(*

**Autonumbered labeled footnotes**

They may be assigned 'autonumber labels' - for instance, [#first]_ and [#second]_. 

--------

.. [#first] a.k.a. first_ 

.. [#second] a.k.a. second_
*)

FUNCTION_BLOCK FB_Libdoc_NamedAutomaticallyNumberedFootnotes
VAR_INPUT
    nVarA : INT;
    nVarB : INT;
END_VAR
VAR_OUTPUT
    nSum : INT;
END_VAR
VAR
END_VAR

END_FUNCTION_BLOCK

(* stored: Version 1.1.0.1, ProductVersion 3.1.4022.17
   POU FB_Libdoc_NamedAutomaticallyNumberedFootnotes: Id {2437e105-852f-45f4-95c4-17ab47dc4611}, SpecialFunc None *)
